Fanuc KAREL source: kd00011.KL

-- PROVISIONAL review KL for V940-1; original PC SHA256 83add3a69ad093fab0dea1d58c9b295b59ff28ce49bd6a10927a676105add631
-- Incomplete behavior may be omitted. Consult companion uncertainty JSON. Do not deploy.
PROGRAM KD00011
%NOLOCKGROUP
VAR
  I : INTEGER
  J : INTEGER
  B : BOOLEAN
  R : REAL
  S : STRING[80]
BEGIN
  -- V9_ZERO_TABLE_METADATA_HINT layout=0001; no indexed target words; source/name/runtime held
  -- UNRESOLVED_PC offsets 5-6; opcodes 15
  -- UNRESOLVED_PC offsets 11-15; opcodes 7F
END KD00011
